(* IEC 61131-3 sources: teller/JD_Teller_LC2_V11/Class/ETVEdge_DigIO_Base, 1 file *)

(* ---- ETVEdge_DigIO_Base.st ---- *)
#include <.\lsl_st_pci.h>

(*!
<Class
	Name               = "ETVEdge_DigIO_Base"
	Revision           = "1.3"
	RealtimeTask       = "false"
	CyclicTask         = "false"
	BackgroundTask     = "false"
	Sigmatek           = "true"
	OSInterface        = "false"
	HighPriority       = "false"
	Automatic          = "false"
	UpdateMode         = "Prescan"
	IconPath           = ".\Class\Tool.ico"
	SharedCommandTable = "true"
	Objectsize         = "(426,120)"
	Comment            = "Class to access digital IOs on Edge Terminals (8xDigIn, 8xDigOut)">
	<Channels>
		<Server Name="Input1" Visualized="true" Initialize="false" WriteProtected="true" Retentive="false"/>
		<Server Name="Input2" Visualized="true" Initialize="false" WriteProtected="true" Retentive="false"/>
		<Server Name="Input3" Visualized="true" Initialize="false" WriteProtected="true" Retentive="false"/>
		<Server Name="Input4" Visualized="true" Initialize="false" WriteProtected="true" Retentive="false"/>
		<Server Name="Input5" Visualized="true" Initialize="false" WriteProtected="true" Retentive="false"/>
		<Server Name="Input6" Visualized="true" Initialize="false" WriteProtected="true" Retentive="false"/>
		<Server Name="Input7" Visualized="true" Initialize="false" WriteProtected="true" Retentive="false"/>
		<Server Name="Input8" Visualized="true" Initialize="false" WriteProtected="true" Retentive="false"/>
		<Server Name="InputByte" Visualized="true" Initialize="false" WriteProtected="false" Retentive="false"/>
		<Server Name="Output1" Visualized="true" Initialize="false" WriteProtected="false" Retentive="false"/>
		<Server Name="Output2" Visualized="true" Initialize="false" WriteProtected="false" Retentive="false"/>
		<Server Name="Output3" Visualized="true" Initialize="false" WriteProtected="false" Retentive="false"/>
		<Server Name="Output4" Visualized="true" Initialize="false" WriteProtected="false" Retentive="false"/>
		<Server Name="Output5" Visualized="true" Initialize="false" WriteProtected="false" Retentive="false"/>
		<Server Name="Output6" Visualized="true" Initialize="false" WriteProtected="false" Retentive="false"/>
		<Server Name="Output7" Visualized="true" Initialize="false" WriteProtected="false" Retentive="false"/>
		<Server Name="Output8" Visualized="true" Initialize="false" WriteProtected="false" Retentive="false"/>
		<Server Name="OutputByte" Visualized="true" Initialize="false" WriteProtected="false" Retentive="false"/>
		<Server Name="State" Visualized="true" Initialize="false" WriteProtected="true" Retentive="false" Comment=" 0..Everything is OK&#13;&#10;-1..Failed to initialize OS-Interface&#13;&#10;-2..IO-Device not available&#13;&#10;-3..Failed to login to HwControl"/>
		<Client Name="To_HwControl" Required="true" Internal="false" Comment="Connect to Client &quot;Control&quot; of &quot;HwControl&quot;-Object"/>
	</Channels>
	<Dependencies>
		<Files>
			<File Path=".\lsl_st_pci.h" Include="true"/>
		</Files>
	</Dependencies>
	<RevDoku>
		<Owner Company="Sigmatek" Author="RamAnd"/>
		<Dokumentation Revision="1.3" Date="14.02.2012" Author="RamAnd" Company="Sigmatek" Description="Outputs are only written to hardware, if they have changed."/>
		<Dokumentation Revision="1.2" Date="27.10.2010" Author="RamAnd" Company="Sigmatek" Description="Added RtPostScan support"/>
		<Dokumentation Revision="1.1" Date="16.07.2010" Author="BleErn" Company="Sigmatek" Description="Servers OutputByte/OutputWord are thread-safe now"/>
		<Dokumentation Revision="1.0" Date="26.02.2010" Author="RamAnd" Company="Sigmatek" Description="Initial version"/>
	</RevDoku>
</Class>
*)
ETVEdge_DigIO_Base : CLASS
	TYPE
	  t_outs : BSINT
	  [
	    1 Supply5VEnable_n,
	    2 LVDSDriverEnable,
	    3 DisplayEnable,
	    4 DisplayBacklightEnable,
	    5 DisplayPowerOn,
	  ];
#pragma pack(push, 1)
	  DigIOs : STRUCT
	    DigOuts : t_outs;
	    DigIns : BSINT
	    [
	    ];
	  END_STRUCT;
#pragma pack(pop)
	END_TYPE
  //Servers:
	State 	: SvrChCmd_DINT;
	Input1 	: SvrCh_DINT;
	Input2 	: SvrCh_DINT;
	Input3 	: SvrCh_DINT;
	Input4 	: SvrCh_DINT;
	Input5 	: SvrCh_DINT;
	Input6 	: SvrCh_DINT;
	Input7 	: SvrCh_DINT;
	Input8 	: SvrCh_DINT;
	Output1 	: SvrCh_DINT;
	Output2 	: SvrCh_DINT;
	Output3 	: SvrCh_DINT;
	Output4 	: SvrCh_DINT;
	Output5 	: SvrCh_DINT;
	Output6 	: SvrCh_DINT;
	Output7 	: SvrCh_DINT;
	Output8 	: SvrCh_DINT;
	InputByte 	: SvrCh_BDINT;
	OutputByte 	: SvrCh_BDINT;
  //Clients:
	To_HwControl 	: CltChCmd_HwControl;
  //Variables:
		pDigs 	: ^DigIOs;
		Power 	: t_outs;
		pSPCIInfo 	: ^LSL_SPCIINFO;
		OutputByteOld : BDINT
		[
		];

		us_FirstScan 	: USINT;
  //Functions:

	FUNCTION VIRTUAL GLOBAL Init;

	FUNCTION VIRTUAL GLOBAL RtWork
		VAR_INPUT
			EAX 	: UDINT;
		END_VAR
		VAR_OUTPUT
			state (EAX) 	: UDINT;
		END_VAR;

	FUNCTION GLOBAL RtPostScan
		VAR_INPUT
			pThis 	: ^DINT;
		END_VAR;

	FUNCTION VIRTUAL GLOBAL Output1::Write
		VAR_INPUT
			input (EAX) 	: DINT;
		END_VAR
		VAR_OUTPUT
			result (EAX) 	: DINT;
		END_VAR;

	FUNCTION VIRTUAL GLOBAL Output2::Write
		VAR_INPUT
			input (EAX) 	: DINT;
		END_VAR
		VAR_OUTPUT
			result (EAX) 	: DINT;
		END_VAR;

	FUNCTION VIRTUAL GLOBAL Output3::Write
		VAR_INPUT
			input (EAX) 	: DINT;
		END_VAR
		VAR_OUTPUT
			result (EAX) 	: DINT;
		END_VAR;

	FUNCTION VIRTUAL GLOBAL Output4::Write
		VAR_INPUT
			input (EAX) 	: DINT;
		END_VAR
		VAR_OUTPUT
			result (EAX) 	: DINT;
		END_VAR;

	FUNCTION VIRTUAL GLOBAL Output5::Write
		VAR_INPUT
			input (EAX) 	: DINT;
		END_VAR
		VAR_OUTPUT
			result (EAX) 	: DINT;
		END_VAR;

	FUNCTION VIRTUAL GLOBAL Output6::Write
		VAR_INPUT
			input (EAX) 	: DINT;
		END_VAR
		VAR_OUTPUT
			result (EAX) 	: DINT;
		END_VAR;

	FUNCTION VIRTUAL GLOBAL Output7::Write
		VAR_INPUT
			input (EAX) 	: DINT;
		END_VAR
		VAR_OUTPUT
			result (EAX) 	: DINT;
		END_VAR;

	FUNCTION VIRTUAL GLOBAL Output8::Write
		VAR_INPUT
			input (EAX) 	: DINT;
		END_VAR
		VAR_OUTPUT
			result (EAX) 	: DINT;
		END_VAR;

	FUNCTION VIRTUAL GLOBAL OutputByte::Write
		VAR_INPUT
			input (EAX) 	: BDINT;
		END_VAR
		VAR_OUTPUT
			result (EAX) 	: BDINT;
		END_VAR;
  //Tables:
	FUNCTION @STD
		VAR_OUTPUT
			ret_code	: CONFSTATES;
		END_VAR;
	FUNCTION GLOBAL TAB @CT_;
END_CLASS;

#pragma usingLtd HwControl

FUNCTION VIRTUAL GLOBAL ETVEdge_DigIO_Base::Init
  VAR
    SigmaTekDevInfo : ^PCICONFDATA;
  END_VAR

  us_FirstScan += 1;

  if us_FirstScan = 10 then
    IF OS_CILGET("PCICONFIG", #pSPCIInfo) =  SYS_ERR_NONE THEN
      SigmaTekDevInfo := SPCIINFO_FINDDEVICE(0x1221,0);
      IF SigmaTekDevInfo <> NIL THEN
        pDigs$pVoid := SPCIINFO_GETADDRESS(SigmaTekDevInfo);
        if pDigs = NIL then
          State := -2;
        else
          // initialisiation OK => we login to HwControl
          if To_HwControl.AddSpecialHW(pThis:=THIS$pVirtualBase, pRtPostScan:=#RtPostScan()) then
            State := -3;
          end_if;
        end_if;
      else
        State := -2;
      end_if;
    else
      State := -1;
    end_if;
  end_if;

END_FUNCTION

FUNCTION VIRTUAL GLOBAL ETVEdge_DigIO_Base::RtWork
	VAR_INPUT
		EAX 	: UDINT;
	END_VAR
	VAR_OUTPUT
		state (EAX) 	: UDINT;
	END_VAR

  if pDigs <> NIL then
    // read inputs
    InputByte  := pDigs^.DigIns;

    // show inputs on servers
    Input1$UDINT := InputByte AND 1;
    Input2$UDINT := (InputByte SHR 1) AND 1;
    Input3$UDINT := (InputByte SHR 2) AND 1;
    Input4$UDINT := (InputByte SHR 3) AND 1;
    Input5$UDINT := (InputByte SHR 4) AND 1;
    Input6$UDINT := (InputByte SHR 5) AND 1;
    Input7$UDINT := (InputByte SHR 6) AND 1;
    Input8$UDINT := (InputByte SHR 7) AND 1;
  end_if;

	state := READY;

END_FUNCTION

FUNCTION VIRTUAL GLOBAL ETVEdge_DigIO_Base::Output1::Write
	VAR_INPUT
		input (EAX) 	: DINT;
	END_VAR
	VAR_OUTPUT
		result (EAX) 	: DINT;
	END_VAR

 	result := input;

  if input then
    OutputByte := OutputByte OR 2#00000001;
    Output1 := 1;
  else
    OutputByte := OutputByte AND 2#11111110;
    Output1 := 0;
  end_if;

END_FUNCTION

FUNCTION VIRTUAL GLOBAL ETVEdge_DigIO_Base::Output2::Write
	VAR_INPUT
		input (EAX) 	: DINT;
	END_VAR
	VAR_OUTPUT
		result (EAX) 	: DINT;
	END_VAR

 	result := input;

  if input then
    OutputByte := OutputByte OR 2#00000010;
    Output2 := 1;
  else
    OutputByte := OutputByte AND 2#11111101;
    Output2 := 0;
  end_if;

END_FUNCTION

FUNCTION VIRTUAL GLOBAL ETVEdge_DigIO_Base::Output3::Write
	VAR_INPUT
		input (EAX) 	: DINT;
	END_VAR
	VAR_OUTPUT
		result (EAX) 	: DINT;
	END_VAR

 	result := input;

  if input then
    OutputByte := OutputByte OR 2#00000100;
    Output3 := 1;
  else
    OutputByte := OutputByte AND 2#11111011;
    Output3 := 0;
  end_if;

END_FUNCTION

FUNCTION VIRTUAL GLOBAL ETVEdge_DigIO_Base::Output4::Write
	VAR_INPUT
		input (EAX) 	: DINT;
	END_VAR
	VAR_OUTPUT
		result (EAX) 	: DINT;
	END_VAR

 	result := input;

  if input then
    OutputByte := OutputByte OR 2#00001000;
    Output4 := 1;
  else
    OutputByte := OutputByte AND 2#11110111;
    Output4 := 0;
  end_if;

END_FUNCTION

FUNCTION VIRTUAL GLOBAL ETVEdge_DigIO_Base::Output5::Write
	VAR_INPUT
		input (EAX) 	: DINT;
	END_VAR
	VAR_OUTPUT
		result (EAX) 	: DINT;
	END_VAR

 	result := input;

  if input then
    OutputByte := OutputByte OR 2#00010000;
    Output5 := 1;
  else
    OutputByte := OutputByte AND 2#11101111;
    Output5 := 0;
  end_if;

END_FUNCTION

FUNCTION VIRTUAL GLOBAL ETVEdge_DigIO_Base::Output6::Write
	VAR_INPUT
		input (EAX) 	: DINT;
	END_VAR
	VAR_OUTPUT
		result (EAX) 	: DINT;
	END_VAR

 	result := input;

  if input then
    OutputByte := OutputByte OR 2#00100000;
    Output6 := 1;
  else
    OutputByte := OutputByte AND 2#11011111;
    Output6 := 0;
  end_if;

END_FUNCTION

FUNCTION VIRTUAL GLOBAL ETVEdge_DigIO_Base::Output7::Write
	VAR_INPUT
		input (EAX) 	: DINT;
	END_VAR
	VAR_OUTPUT
		result (EAX) 	: DINT;
	END_VAR

 	result := input;

  if input then
    OutputByte := OutputByte OR 2#01000000;
    Output7 := 1;
  else
    OutputByte := OutputByte AND 2#10111111;
    Output7 := 0;
  end_if;

END_FUNCTION

FUNCTION VIRTUAL GLOBAL ETVEdge_DigIO_Base::Output8::Write
	VAR_INPUT
		input (EAX) 	: DINT;
	END_VAR
	VAR_OUTPUT
		result (EAX) 	: DINT;
	END_VAR

 	result := input;

  if input then
    OutputByte := OutputByte OR 2#10000000;
    Output8 := 1;
  else
    OutputByte := OutputByte AND 2#01111111;
    Output8 := 0;
  end_if;

END_FUNCTION

FUNCTION VIRTUAL GLOBAL ETVEdge_DigIO_Base::OutputByte::Write
	VAR_INPUT
		input (EAX) 	: BDINT;
	END_VAR
	VAR_OUTPUT
		result (EAX) 	: BDINT;
	END_VAR

	result := OutputByte := input;

  // show outputs on servers
  Output1$UDINT := input AND 1;
  Output2$UDINT := (input SHR 1) AND 1;
  Output3$UDINT := (input SHR 2) AND 1;
  Output4$UDINT := (input SHR 3) AND 1;
  Output5$UDINT := (input SHR 4) AND 1;
  Output6$UDINT := (input SHR 5) AND 1;
  Output7$UDINT := (input SHR 6) AND 1;
  Output8$UDINT := (input SHR 7) AND 1;

END_FUNCTION

FUNCTION GLOBAL ETVEdge_DigIO_Base::RtPostScan
	VAR_INPUT
		pThis 	: ^DINT;
	END_VAR

  // we restore our this pointer, because this method is called from hwcontrol
  this$^DINT := pThis;

  if pDigs <> NIL then
    // if they have changed, write the outputs
    IF OutputByte <> OutputByteOld THEN
      pDigs^.DigOuts := OutputByteOld$USINT := OutputByte$usint;
    END_IF;
  end_if;

END_FUNCTION
